(* IEC 61131-3 sources: trust-platform/examples/tutorials, 9 files *)

(* ---- 01_hello_counter.st ---- *)
PROGRAM HelloCounter
VAR
    Enable : BOOL := TRUE;
    ResetCmd : BOOL := FALSE;
    Increment : DINT := 1;
    Count : DINT := 0;
END_VAR

IF ResetCmd THEN
    Count := 0;
ELSIF Enable THEN
    Count := Count + Increment;
END_IF;
END_PROGRAM

(* ---- 02_blinker.st ---- *)
PROGRAM Blinker
VAR
    Enable : BOOL := TRUE;
    Lamp : BOOL := FALSE;
    PulsePeriod : TIME := T#250ms;
    TimerEnable : BOOL := TRUE;
    BlinkTimer : TON;
END_VAR

BlinkTimer(IN := TimerEnable, PT := PulsePeriod);

IF NOT Enable THEN
    Lamp := FALSE;
    TimerEnable := FALSE;
ELSIF BlinkTimer.Q THEN
    Lamp := NOT Lamp;
    TimerEnable := FALSE;
ELSE
    TimerEnable := TRUE;
END_IF;
END_PROGRAM

(* ---- 03_traffic_light.st ---- *)
PROGRAM TrafficLight
VAR
    Phase : INT := 0;
    PhasePeriod : TIME := T#500ms;
    PhaseTimerEnable : BOOL := TRUE;
    PhaseTimer : TON;
    Red : BOOL := TRUE;
    Yellow : BOOL := FALSE;
    Green : BOOL := FALSE;
END_VAR

PhaseTimer(IN := PhaseTimerEnable, PT := PhasePeriod);

CASE Phase OF
    0:
        Red := TRUE;
        Yellow := FALSE;
        Green := FALSE;
    1:
        Red := TRUE;
        Yellow := TRUE;
        Green := FALSE;
    2:
        Red := FALSE;
        Yellow := FALSE;
        Green := TRUE;
    3:
        Red := FALSE;
        Yellow := TRUE;
        Green := FALSE;
END_CASE;

IF PhaseTimer.Q THEN
    CASE Phase OF
        0:
            Phase := 1;
        1:
            Phase := 2;
        2:
            Phase := 3;
        3:
            Phase := 0;
    END_CASE;
    PhaseTimerEnable := FALSE;
ELSE
    PhaseTimerEnable := TRUE;
END_IF;
END_PROGRAM

(* ---- 04_tank_level.st ---- *)
PROGRAM TankLevel
VAR
    InletValveCmd : BOOL := FALSE;
    OutletValveCmd : BOOL := TRUE;
    LevelPercent : REAL := 45.0;
    LowSetpoint : REAL := 30.0;
    HighSetpoint : REAL := 70.0;
END_VAR

IF LevelPercent <= LowSetpoint THEN
    InletValveCmd := TRUE;
    OutletValveCmd := FALSE;
ELSIF LevelPercent >= HighSetpoint THEN
    InletValveCmd := FALSE;
    OutletValveCmd := TRUE;
END_IF;

IF InletValveCmd THEN
    LevelPercent := LevelPercent + 2.5;
END_IF;

IF OutletValveCmd THEN
    LevelPercent := LevelPercent - 1.5;
END_IF;
END_PROGRAM

(* ---- 05_motor_starter.st ---- *)
PROGRAM MotorStarter
VAR
    StartPb : BOOL := FALSE;
    StopPb : BOOL := FALSE;
    OverloadTrip : BOOL := FALSE;
    MotorRun : BOOL := FALSE;
    SealInContact : BOOL := FALSE;
END_VAR

IF StopPb OR OverloadTrip THEN
    MotorRun := FALSE;
ELSIF StartPb OR SealInContact THEN
    MotorRun := TRUE;
END_IF;

SealInContact := MotorRun;
END_PROGRAM

(* ---- 06_recipe_manager.st ---- *)
PROGRAM RecipeManager
VAR
    SelectedRecipe : INT := 1;
    ApplySelection : BOOL := TRUE;
    ActiveTargetTemperature : REAL := 0.0;
    ActiveMixTime : TIME := T#0s;
    ActiveBatchSize : INT := 0;
END_VAR

IF ApplySelection THEN
    CASE SelectedRecipe OF
        1:
            ActiveTargetTemperature := 65.0;
            ActiveMixTime := T#30s;
            ActiveBatchSize := 10;
        2:
            ActiveTargetTemperature := 72.5;
            ActiveMixTime := T#45s;
            ActiveBatchSize := 14;
        3:
            ActiveTargetTemperature := 80.0;
            ActiveMixTime := T#60s;
            ActiveBatchSize := 18;
        ELSE
            ActiveTargetTemperature := 60.0;
            ActiveMixTime := T#20s;
            ActiveBatchSize := 8;
    END_CASE;
END_IF;
END_PROGRAM

(* ---- 07_pid_loop.st ---- *)
PROGRAM PidLoop
VAR
    Setpoint : REAL := 50.0;
    ProcessValue : REAL := 40.0;
    Kp : REAL := 1.2;
    Ki : REAL := 0.1;
    Kd : REAL := 0.05;
    SampleTime : REAL := 0.1;
    IntegralTerm : REAL := 0.0;
    PreviousError : REAL := 0.0;
    ErrorValue : REAL := 0.0;
    Derivative : REAL := 0.0;
    ControlOutput : REAL := 0.0;
END_VAR

ErrorValue := Setpoint - ProcessValue;
IntegralTerm := IntegralTerm + (ErrorValue * Ki * SampleTime);
Derivative := (ErrorValue - PreviousError) / SampleTime;
ControlOutput := (Kp * ErrorValue) + IntegralTerm + (Kd * Derivative);
PreviousError := ErrorValue;
ProcessValue := ProcessValue + (ControlOutput * 0.02);
END_PROGRAM

(* ---- 08_conveyor_system.st ---- *)
PROGRAM ConveyorSystem
VAR
    StartCmd : BOOL := FALSE;
    StopCmd : BOOL := FALSE;
    JamSensor : BOOL := FALSE;
    PartAtEntry : BOOL := FALSE;
    PartAtExit : BOOL := FALSE;
    ConveyorRun : BOOL := FALSE;
    RejectGate : BOOL := FALSE;
    PartCounter : DINT := 0;
END_VAR

IF StopCmd OR JamSensor THEN
    ConveyorRun := FALSE;
ELSIF StartCmd THEN
    ConveyorRun := TRUE;
END_IF;

IF ConveyorRun AND PartAtEntry THEN
    RejectGate := FALSE;
END_IF;

IF ConveyorRun AND PartAtExit THEN
    PartCounter := PartCounter + 1;
END_IF;

IF JamSensor THEN
    RejectGate := TRUE;
END_IF;
END_PROGRAM

(* ---- 09_simulation_coupling.st ---- *)
PROGRAM SimulationCouplingDemo
VAR
    TankLevelRaw : WORD;
    HighLevelAlarm : BOOL;
END_VAR

HighLevelAlarm := WORD_TO_UINT(TankLevelRaw) >= 500;
END_PROGRAM

CONFIGURATION SimulationCouplingConfig
TASK Cycle (INTERVAL := T#100ms, PRIORITY := 1);
PROGRAM P1 WITH Cycle : SimulationCouplingDemo;
VAR_CONFIG
    P1.TankLevelRaw AT %IW0 : WORD;
    P1.HighLevelAlarm AT %QX0.0 : BOOL;
END_VAR
END_CONFIGURATION
